// TwinCAT 3 PLC project FoE
// ProgramVersion: 3.1.4023.0
// libraries:
//   Tc2_EtherCAT, * (Beckhoff Automation GmbH)
//   Tc2_Standard, * (Beckhoff Automation GmbH)
//   Tc2_System, * (Beckhoff Automation GmbH)
//   Tc3_Module, * (Beckhoff Automation GmbH)
// project tree:
//   / PlcTask.TcTTO
//   POUs/ MAIN.TcPOU
// real-time tasks:
//   TASK PlcTask: cycle T#10ms, priority 20, ADS port 350
// I/O:
//   DEVICE Device 2 (EtherCAT), AmsNetId 192.168.18.191.3.1
//     Box 1 (LAN9255_EtherCAT_Slave) [LAN9255_EtherCAT_Slave]

CONFIGURATION FoE
    RESOURCE PLC ON TwinCAT3
        TASK PlcTask(INTERVAL := T#10ms, PRIORITY := 20);
        PROGRAM MAIN WITH PlcTask : MAIN;
    END_RESOURCE
END_CONFIGURATION

// ---- POUs/MAIN.TcPOU
PROGRAM MAIN
VAR
	
    fbDownload : FB_EcFoeLoad ;
		
	dwPass	: DWORD := 287454020; // 0x11223344
	sNetId     : T_AmsNetId := '192.168.18.191.3.1' ;
    nSlaveAddr : UINT := 1001;  
	eMode      : E_EcFoeMode := eFoeMode_Write;
	sPathName : STRING := 'D:\LAN9255Updated.bin';
	
    bLoad      : BOOL;
    bBusy      : BOOL;
    bError     : BOOL;
    nErrID     : UDINT;
    nBytesWritten : UDINT;
    nPercent      : UDINT;
END_VAR

fbDownload( bExecute := bLoad,
		sNetId  := sNetId,
		nSlaveAddr := nSlaveAddr,
		dwPass  := dwPass,
		sPathName  := sPathName, 
        bBusy => bBusy,
        bError => bError,
        nErrId => nErrID,
        cbLoad => nBytesWritten,
        nProgress => nPercent );

END_PROGRAM
